Fanuc KAREL source: KA00013.KL

PROGRAM KA00013
%NOLOCKGROUP
VAR
  SRC: REAL
  DST: INTEGER
BEGIN
  SRC = 2.0
  DST = SRC
END KA00013
